TYPE ST_PolarIIChamber_NozzlePortServiceStatus :
STRUCT
	Nozzle : ARRAY[1..3] OF ST_PolarIIChamber_PortNozzleSupplyServiceStatus;
	DrainSelect1 : ST_ServiceStatus;
	DrainSelect2 : ST_ServiceStatus;
	DrainSelect3 : ST_ServiceStatus;
END_STRUCT
END_TYPE

(* stored: Version 1.1.0.1, ProductVersion 3.1.4026.18
   DUT ST_PolarIIChamber_NozzlePortServiceStatus: Id {14000000-0000-0000-0000-000000000057} *)
